(* IEC 61131-3 sources: plc-iiot-stack/src/POUs/Iiot/FB_MqttAlarms, 10 files *)

(* ---- FB_MqttAlarms.decl.st ---- *)
// Назначение: публикация событий тревог (data_schema 4) в <prefix>/<device>/alarm/<suffix>, QoS 1, retain:
//             {schema_version, ts, id, code, priority, state, prev_state, reason}. Состояние тревоги — по
//             словам устройства (wAlmActive, wAlmUnack, wAlmShelved, режим OutOfService); событие — смена
//             состояния с прошлой публикации, причина — по переходу (F_IiotAlarmReason). После каждого
//             рождения узла (xReady) публикуются все тревоги: не менявшаяся — повтором последней
//             публикации с её ts (в InfluxDB та же точка, не новое срабатывание), изменившаяся без связи —
//             событием, ещё не публиковавшаяся с запуска ПЛК — снимком (prev_state = state). Переходы между
//             двумя публикациями сливаются в один; точные события ST_AlarmEvent во флагмане даёт
//             PL.I_AlarmSink (docs/plc_mqtt.md).
// Автор:      kr0nsch
// Версия:     0.1.1
// Документ:   docs/plc_mqtt.md, раздел «Тревоги»
FUNCTION_BLOCK FB_MqttAlarms
VAR_INPUT
    xEnable : BOOL;
    xReady : BOOL;                                        // связь есть и рождение опубликовано
    itfClient : I_MqttClient;
    uliTs_ms : ULINT;                                     // время UTC, мс (поле ts)
    sTopicPrefix : STRING(GVL_Const.IIOT_PREFIX_LEN);     // site/area/unit
    uiMaxPerCycle : UINT := GVL_Const.ALARMS_MAX_PER_CYCLE;
END_VAR
VAR_IN_OUT
    aAlarms : ARRAY[*] OF ST_IiotAlarm;
    aWords : ARRAY[*] OF ST_IiotAlarmWords;               // строки — ST_IiotAlarmCfg.diWords
END_VAR
VAR_OUTPUT
    udiPublished : UDINT;
    udiFailed : UDINT;
    udiDropped : UDINT;
    udiEvents : UDINT;          // опубликовано событий (без снимков)
    uiPending : UINT;
END_VAR
VAR
    fbJson : FB_JsonBuilder;
    sTopic : STRING(GVL_Const.MQTT_TOPIC_LEN);
    diCursor : DINT;
END_VAR

(* ---- FB_MqttAlarms.impl.st ---- *)
// Состояние каждой тревоги — каждый вызов (видно и без связи)
UpdateStates(aAlarmTable := aAlarms, aWordTable := aWords);

IF NOT xEnable OR NOT xReady OR itfClient = 0 OR NOT F_IiotClockValid(uliTs_ms := uliTs_ms) THEN
    ResetSent(aAlarmTable := aAlarms);
    RETURN;
END_IF
IF NOT itfClient.IsConnected() THEN
    ResetSent(aAlarmTable := aAlarms);
    RETURN;
END_IF
PublishDue(aAlarmTable := aAlarms);

(* ---- PublishAlarm.method.decl.st ---- *)
// Опубликовать тревогу. TRUE — обработана (опубликована или пропущена). Что публикуется:
// - событие: состояние изменилось с прошлой публикации (в том числе пока связи не было) — ts сейчас;
// - повтор после переподключения: состояние не менялось — последняя публикация с её ts и prev_state
//   (в InfluxDB та же точка: активная тревога не считается новым срабатыванием);
// - снимок: с запуска ПЛК тревога не публиковалась — prev_state = state, ts сейчас.
METHOD PRIVATE PublishAlarm : BOOL
VAR_IN_OUT
    stAlarm : ST_IiotAlarm;
END_VAR
VAR
    ePrev : E_IiotAlarmState;
    uliTs : ULINT;
    xEvent : BOOL;
    sCode : STRING(GVL_Const.IIOT_TEXT_LEN);
    sPriority : STRING(GVL_Const.IIOT_TEXT_LEN);
    sPath : STRING(GVL_Const.MQTT_TOPIC_LEN);
END_VAR

(* ---- PublishAlarm.method.impl.st ---- *)
uliTs := uliTs_ms;
IF stAlarm.xSent OR (stAlarm.uliEventTs_ms > 0 AND stAlarm.eState <> stAlarm.eLastState) THEN
    xEvent := TRUE;                     // событие: в том числе переход, случившийся без связи
    ePrev := stAlarm.eLastState;
ELSIF stAlarm.uliEventTs_ms > 0 THEN
    xEvent := FALSE;                    // повтор последней публикации после переподключения
    ePrev := stAlarm.eEventPrev;
    uliTs := stAlarm.uliEventTs_ms;
ELSE
    xEvent := FALSE;                    // снимок: с запуска ПЛК не публиковалась
    ePrev := stAlarm.eState;
END_IF
sPriority := F_IiotAlarmPriorityText(ePriority := stAlarm.stCfg.ePriority);
sCode := CONCAT(CONCAT(stAlarm.stCfg.sDevice, '.'), stAlarm.stCfg.sSuffix);
sPath := CONCAT(CONCAT(stAlarm.stCfg.sDevice, GVL_Const.TOPIC_SEPARATOR), GVL_Const.TOPIC_ALARM_LEVEL);
sPath := CONCAT(CONCAT(sPath, GVL_Const.TOPIC_SEPARATOR), stAlarm.stCfg.sSuffix);
sTopic := F_IiotTopic(sPrefix := sTopicPrefix, sPath := sPath);
fbJson.Begin();
fbJson.AddString(sKey := 'schema_version', sValue := GVL_Const.IIOT_SCHEMA_VERSION);
fbJson.AddInt(sKey := 'ts', liValue := ULINT_TO_LINT(uliTs));
fbJson.AddInt(sKey := 'id', liValue := UDINT_TO_LINT(stAlarm.stCfg.udiId));
fbJson.AddString(sKey := 'code', sValue := sCode);
fbJson.AddString(sKey := 'priority', sValue := sPriority);
fbJson.AddString(sKey := 'state', sValue := F_IiotAlarmStateText(eState := stAlarm.eState));
fbJson.AddString(sKey := 'prev_state', sValue := F_IiotAlarmStateText(eState := ePrev));
fbJson.AddString(sKey := 'reason',
                 sValue := F_IiotAlarmReasonText(eReason := F_IiotAlarmReason(ePrev := ePrev, eNew := stAlarm.eState)));

IF NOT fbJson.Finish() OR LEN(sTopic) = 0 OR LEN(sPriority) = 0 THEN
    udiDropped := udiDropped + 1;
ELSIF itfClient.Publish(sTopic := sTopic, eQos := E_MqttQos.AtLeastOnce, xRetain := TRUE,
                        sPayload := fbJson.sJson) THEN
    udiPublished := udiPublished + 1;
    IF xEvent THEN
        udiEvents := udiEvents + 1;
    END_IF
ELSE
    udiFailed := udiFailed + 1;
    RETURN;
END_IF
stAlarm.eLastState := stAlarm.eState;
stAlarm.eEventPrev := ePrev;
stAlarm.uliEventTs_ms := uliTs;
stAlarm.xSent := TRUE;
PublishAlarm := TRUE;

(* ---- PublishDue.method.decl.st ---- *)
// Обход тревог по кругу: не опубликована с подключения (снимок или повтор) или состояние изменилось (событие).
METHOD PRIVATE PublishDue
VAR_IN_OUT
    aAlarmTable : ARRAY[*] OF ST_IiotAlarm;
END_VAR
VAR
    diLo : DINT;
    diTotal : DINT;
    diStep : DINT;
    diIdx : DINT;
    diNextCursor : DINT;
    uiBudget : UINT;
    xBlocked : BOOL;
END_VAR

(* ---- PublishDue.method.impl.st ---- *)
diLo := LOWER_BOUND(aAlarmTable, 1);
diTotal := UPPER_BOUND(aAlarmTable, 1) - diLo + 1;
uiPending := 0;
IF diTotal <= 0 THEN
    RETURN;
END_IF
IF diCursor < 0 OR diCursor >= diTotal THEN
    diCursor := 0;
END_IF
uiBudget := MAX(uiMaxPerCycle, 1);
diNextCursor := -1;
FOR diStep := 0 TO diTotal - 1 DO
    diIdx := diLo + (diCursor + diStep) MOD diTotal;
    IF NOT aAlarmTable[diIdx].xSent OR aAlarmTable[diIdx].eState <> aAlarmTable[diIdx].eLastState THEN
        IF uiBudget > 0 AND NOT xBlocked THEN
            IF PublishAlarm(stAlarm := aAlarmTable[diIdx]) THEN
                uiBudget := uiBudget - 1;
            ELSE
                xBlocked := TRUE;
            END_IF
        END_IF
        IF NOT aAlarmTable[diIdx].xSent OR aAlarmTable[diIdx].eState <> aAlarmTable[diIdx].eLastState THEN
            uiPending := uiPending + 1;
            IF diNextCursor < 0 THEN
                diNextCursor := diIdx - diLo;
            END_IF
        END_IF
    END_IF
END_FOR
IF diNextCursor >= 0 THEN
    diCursor := diNextCursor;
END_IF

(* ---- ResetSent.method.decl.st ---- *)
// Связи нет: после рождения узла публикуются все тревоги (повтор, событие или снимок — PublishAlarm).
METHOD PRIVATE ResetSent
VAR_IN_OUT
    aAlarmTable : ARRAY[*] OF ST_IiotAlarm;
END_VAR
VAR
    diIdx : DINT;
END_VAR

(* ---- ResetSent.method.impl.st ---- *)
FOR diIdx := LOWER_BOUND(aAlarmTable, 1) TO UPPER_BOUND(aAlarmTable, 1) DO
    aAlarmTable[diIdx].xSent := FALSE;
END_FOR
uiPending := 0;

(* ---- UpdateStates.method.decl.st ---- *)
// Состояние каждой тревоги по словам её устройства; строка слов вне таблицы — тревога в норме.
METHOD PRIVATE UpdateStates
VAR_IN_OUT
    aAlarmTable : ARRAY[*] OF ST_IiotAlarm;
    aWordTable : ARRAY[*] OF ST_IiotAlarmWords;
END_VAR
VAR
    diIdx : DINT;
    diWords : DINT;
END_VAR

(* ---- UpdateStates.method.impl.st ---- *)
FOR diIdx := LOWER_BOUND(aAlarmTable, 1) TO UPPER_BOUND(aAlarmTable, 1) DO
    diWords := aAlarmTable[diIdx].stCfg.diWords;
    IF diWords >= LOWER_BOUND(aWordTable, 1) AND diWords <= UPPER_BOUND(aWordTable, 1) THEN
        aAlarmTable[diIdx].eState := F_IiotAlarmStateOf(stWords := aWordTable[diWords],
                                                        uiSlot := aAlarmTable[diIdx].stCfg.uiSlot);
    ELSE
        aAlarmTable[diIdx].eState := E_IiotAlarmState.Normal;
    END_IF
END_FOR
